// Target for the ADS RPC tests: AddNumbers is callable through ADS by symbol name.
FUNCTION_BLOCK T_RpcTarget
VAR
  _lastSum : DINT;
END_VAR

{attribute 'TcRpcEnable'}
METHOD AddNumbers : DINT
VAR_INPUT
  a : DINT;
  b : DINT;
END_VAR
AddNumbers := a + b;
_lastSum := AddNumbers;
END_METHOD

PROPERTY LastSum : DINT
GET
LastSum := _lastSum;
END_GET
END_PROPERTY

END_FUNCTION_BLOCK

(* stored: Version 1.1.0.1, ProductVersion 3.1.4026.22
   POU T_RpcTarget: Id {44ec3c53-cc59-420b-a59a-70bb63636348}, SpecialFunc None
   Method AddNumbers: Id {abc64f41-a75c-45a0-a069-9cfd11f7948b}
   Property LastSum: Id {a0ee6918-dde5-4689-ab8e-17fd5559396d}
   Get Get: Id {a8e4f882-08f6-4e60-b986-8730919faf14} *)
